TYPE E_userGroup :
(
	Group1:=1,
	Group2:=2,
	Group3:=3,
	Group4:=4
);
END_TYPE

(* stored: Version 1.1.0.1, ProductVersion 3.1.4024.13
   DUT E_userGroup: Id {acdb8d99-e806-4262-9edf-ab1b53b06e04} *)
